(* IEC 61131-3 sources: codesys-to-astra/src/POUs/F_C2aBefore, 2 files *)

(* ---- F_C2aBefore.decl.st ---- *)
// Назначение: замена OSU.Before (OwenStringUtils v3.0, с. 15): фрагмент sSource до первого вхождения
//             sPostfix; не найдено — пустая строка.
// Автор:      kr0nsch
// Версия:     0.1.0
// Документ:   docs/LIBMAP.md
FUNCTION F_C2aBefore : STRING(255)
VAR_INPUT
    sSource : STRING(255);  // исходная строка
    sPostfix : STRING(255); // подстрока
END_VAR
VAR
    iPos : INT;             // позиция вхождения (с 1) или 0
END_VAR

(* ---- F_C2aBefore.impl.st ---- *)
iPos := FIND(sSource, sPostfix);
IF iPos > 0 AND LEN(sPostfix) > 0 THEN
    F_C2aBefore := LEFT(sSource, iPos - 1);
ELSE
    F_C2aBefore := '';
END_IF
